(* PLC project g_transformer_protect_bomb, Anonymous Benchmark Suite 1.0 *)
(* stored: creationDateTime 2026-07-09T00:00:00 *)

PROGRAM g_transformer_protect_bomb
  VAR_INPUT
    energize_cmd : BOOL;
    oil_temp_high : BOOL;
    lockout : BOOL;
    maint : BOOL;
  END_VAR
  VAR_OUTPUT
    transformer_on : BOOL;
    trip : BOOL;
  END_VAR

(* LD diagram, written out as Structured Text *)
transformer_on := (NOT oil_temp_high OR oil_temp_high AND maint) AND energize_cmd AND NOT lockout;
trip := oil_temp_high;
END_PROGRAM

CONFIGURATION Config0
  RESOURCE Res0 ON PLC
    TASK tcyclic(INTERVAL := T#10ms, PRIORITY := 0);
    PROGRAM inst0 WITH tcyclic : g_transformer_protect_bomb;
  END_RESOURCE
END_CONFIGURATION
